(* IEC 61131-3 sources: JingjiangMoonbox/Application/Application/任务列表/Main_Task/GNS_MAP/STRUCT/ENUM, 4 files *)

(* ---- stEnumAxisId.st ---- *)
(*@CES
Name=stEnumAxisId
Type=Gvl
TypeGuid=2db5746d-d284-4425-9f7f-2663a34b0ebc
Guid=4f97fc19-ca37-4da0-90af-5aea95a45e3f
HasDeclaration=True
HasImplementation=False
*)
{DECLARATION}
//{attribute 'qualified_only'}
{attribute 'strict'}
TYPE stEnumAxisId :(
	AXISID_INVALID:=-1,
	AXISID_RESERVED,
	(*不能随意调整@start*)
	AXISID_1U:=1,
	AXISID_2U,
	AXISID_3U,
	AXISID_4U,
	AXISID_5U,
	AXISID_6U,
	AXISID_7U,
	AXISID_8U,
	AXISID_9U,
	AXISID_10U,
	AXISID_11U,
	AXISID_12U,
	AXISID_13U,
	AXISID_14U,
	AXISID_15U,
	(*不能随意调整@end*)
	AXISID_UWA,(*放料A*)
	AXISID_UWB,
	AXISID_RWA,
	AXISID_RWB,
	AXISID_IF,(*放牵*)
	AXISID_OF,
	AXISID_UWA_II,
	AXISID_UWB_II,
	AXISID_RWA_II,
	AXISID_RWB_II,
	AXISID_IF_II,
	AXISID_OF_II,
	AXISID_CENTER(*中心辊*)
);
END_TYPE

{IMPLEMENTATION}

(* ---- stEnumFuncId.st ---- *)
(*@CES
Name=stEnumFuncId
Type=Gvl
TypeGuid=2db5746d-d284-4425-9f7f-2663a34b0ebc
Guid=977dc716-2507-48a6-a21c-666c8469de7d
HasDeclaration=True
HasImplementation=False
*)
{DECLARATION}
//{attribute 'qualified_only'}
{attribute 'strict'}
TYPE stEnumFuncId :((*色组驱动器的功能id*)
	FUNCID_NULL :=-1,(*无功能*)
	FUNCID_RESERVED,(*占位*)
	(*站的功能*)
	FUNCID_CONTROL,(*控制功能@目前架构应该是月光系列*)
	FUNCID_PRNROLLER,(*版辊*)
	FUNCID_NETROLLER,(*网辊*)
	FUNCID_BOTTOMROLLER,(*底辊*)
	FUNCID_PRNROLLER_PRESSURE_M,(*版辊压力|操作侧*)
	FUNCID_PRNROLLER_PRESSURE_G,
	FUNCID_NETROLLER_PRESSURE_M,(*网辊压力|操作侧*)
	FUNCID_NETROLLER_PRESSURE_G,
	FUNCID_HORZ,(*横向*)
	(*龙门功能id@*)
	FUNCID_PRNROLLER_GANTRY,(*印刷辊龙门*)
	FUNCID_NETROLLER_GANTRY(*网纹辊龙门*)
);
END_TYPE

{IMPLEMENTATION}

(* ---- stEnumMoveType.st ---- *)
(*@CES
Name=stEnumMoveType
Type=Gvl
TypeGuid=2db5746d-d284-4425-9f7f-2663a34b0ebc
Guid=686aa444-d3fe-4889-be0c-cd0099a56b1b
HasDeclaration=True
HasImplementation=False
*)
{DECLARATION}
//{attribute 'qualified_only'}
{attribute 'strict'}
TYPE stEnumMoveType :((*运动类型*)
	MOVETYPE_NULL :=0,(*不运动*)
	MOVETYPE_TRAP ,(*点位运动*)
	MOVETYPE_GANTRY,(*龙门运动*)
	MOVETYPE_ROTARY,(*旋转电机*)
	MOVETYPE_ROTARY_SUPERPOS(*旋转电机-叠加位置*)
);
END_TYPE
{IMPLEMENTATION}

(* ---- stEuumMachineryType.st ---- *)
(*@CES
Name=stEuumMachineryType
Type=Gvl
TypeGuid=2db5746d-d284-4425-9f7f-2663a34b0ebc
Guid=aab11485-0b5d-4c95-bba7-862ff1a86d0f
HasDeclaration=True
HasImplementation=False
*)
{DECLARATION}
//{attribute 'qualified_only'}
{attribute 'strict'}
TYPE stEuumMachineryType :((*机器类型*)
	MACHINERYTYPE_ROTOGRAVE,(*凹版印刷机*)
	MACHINERYTYPE_FELXO_INLINE,(*机组式柔印@套色叠加轴在网辊*)
	MACHINERYTYPE_FELXO_INLINE_ONEBOTOMROLLER,(*机组式柔印@单底辊(套色叠加轴是需要在底辊上)*)
	MACHINERYTYPE_FELXO_CL,(*卫星式柔印*)
	MACHINERYTYPE_OFFSET(*胶印机*)
);
END_TYPE
{IMPLEMENTATION}
